(* Logix 5000 project; controller R400_500_XLS vendor 1 type 14 code 216 rev 31.11; software revision 31.01; part 13 of 32 *)
(* tags used below, declared in another part *)
   Alarm : SINT;   // Wait 3 seconds
   AlarmMuted : BOOL;
   Chem_Pump : UDT_CHEM_PUMP[4];   // Chemical Pump flow rate
   ChPumpRunningTime : REAL;
   Inj_Cond : SINT;   // Conductivity injection based steps
   Inj_Time : SINT;   // Time based chemical injection steps
   M : DINT[5];   // Memory Bits
   NeutralizantPump : SINT;
   NeutralizationInjTime : DINT;
   NeutralizationRecircTime : DINT;
   OneShot : DINT[1];
   Run : DINT;
   Service : DINT[2];   // Unused Service Mode Memory Bit
   Supervisor : DINT;
   Tmr : TIMER[107];
   VolumeInjected_ML : REAL;
   VolumeNeutralizer : REAL;
   washerMode : SINT;   // Washer Mode Flag 0 -> Ready; 1 -> Supervisor; 2 -> Service; 3 -> Run.
   WshExcBuffer : UDT_WASH;
   Current_Screen : DINT;
   Doors_Check : DINT;
   NumInput : UDT_NUMERIC_INPUT[65];   // Numeric input
   NumInputReal : UDT_NUMERIC_INPUT_REAL[17];
   Q_Chm_1 : BOOL;   // Chemical pump #1
   Q_Chm_2 : BOOL;   // Chemical pump #2
   Q_Chm_3 : BOOL;   // Chemical pump #3
   Q_Chm_4 : BOOL;   // Chemical pump #4
   Screen_Ctrl : DINT;   // PLC Screen Request
   SelChemNeutralizer : UDT_SELECTOR[5];
   SelChemNeutralizerESign : UDT_SELECTOR[5];
   Selector : UDT_SELECTOR[25];   // Piloted list selector
   Tpb : DINT[11];
   udtAudibleAlarmMode : UDT_SELECTOR;
   Unit : Hrdwre;   // Unit Configuration
(* MainProgram, continued *)

ROUTINE SPV_18_AUDIBLE_ALARM_OP_MODE   (* ladder *)
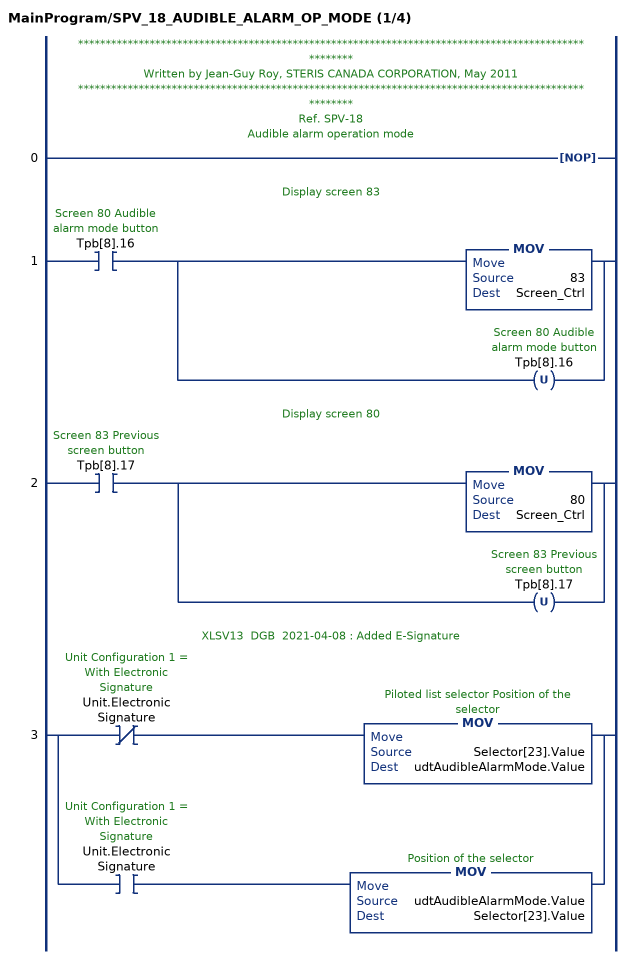
   // ****************************************************************************************************
   // Written by Jean-Guy Roy, STERIS CANADA CORPORATION, May 2011
   // ****************************************************************************************************
   // Ref. SPV-18
   // Audible alarm operation mode
   0: NOP();
   // Display screen 83
   1: XIC(Tpb[8].16)[MOV(83,Screen_Ctrl) ,OTU(Tpb[8].16) ];
   // Display screen 80
   2: XIC(Tpb[8].17)[MOV(80,Screen_Ctrl) ,OTU(Tpb[8].17) ];
   // XLSV13  DGB  2021-04-08 : Added E-Signature
   3: [XIO(Unit.ElectronicSignature) MOV(Selector[23].Value,udtAudibleAlarmMode.Value) ,XIC(Unit.ElectronicSignature) MOV(udtAudibleAlarmMode.Value,Selector[23].Value) ];
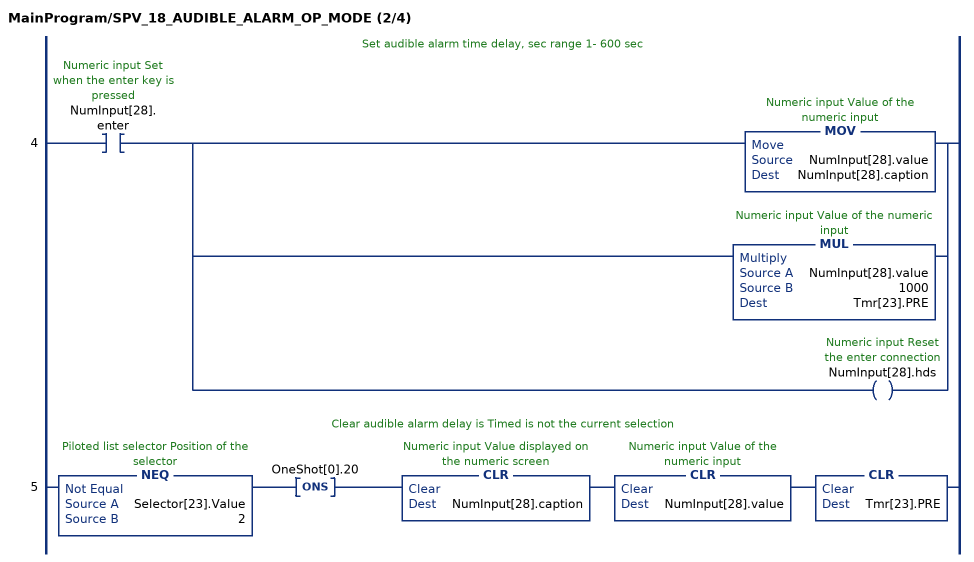
   // Set audible alarm time delay, sec range 1- 600 sec
   4: XIC(NumInput[28].enter)[MOV(NumInput[28].value,NumInput[28].caption) ,MUL(NumInput[28].value,1000,Tmr[23].PRE) ,OTE(NumInput[28].hds) ];
   // Clear audible alarm delay is Timed is not the current selection
   5: NEQ(Selector[23].Value,2)ONS(OneShot[0].20)CLR(NumInput[28].caption)CLR(NumInput[28].value)CLR(Tmr[23].PRE);
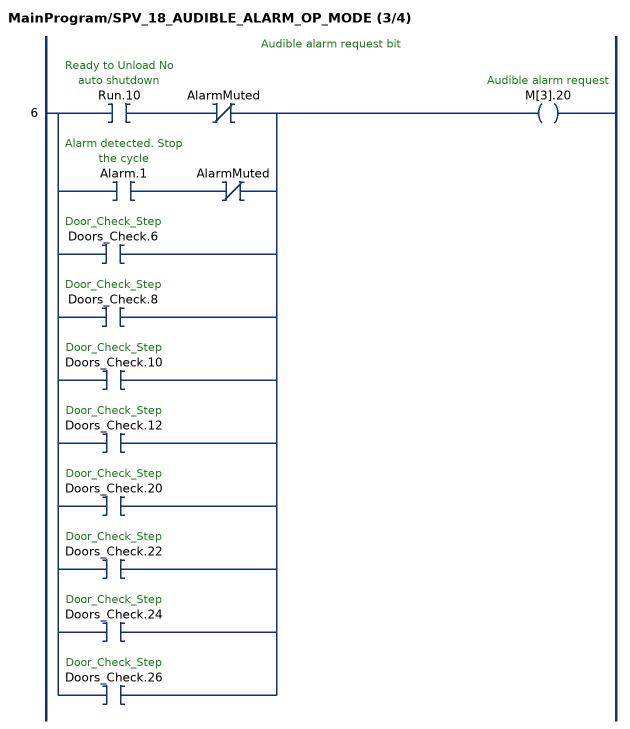
   // Audible alarm request bit
   6: [XIC(Run.10) XIO(AlarmMuted) ,XIC(Alarm.1) XIO(AlarmMuted) ,XIC(Doors_Check.6) ,XIC(Doors_Check.8) ,XIC(Doors_Check.10) ,XIC(Doors_Check.12) ,XIC(Doors_Check.20) ,XIC(Doors_Check.22) ,XIC(Doors_Check.24) ,XIC(Doors_Check.26) ]OTE(M[3].20);
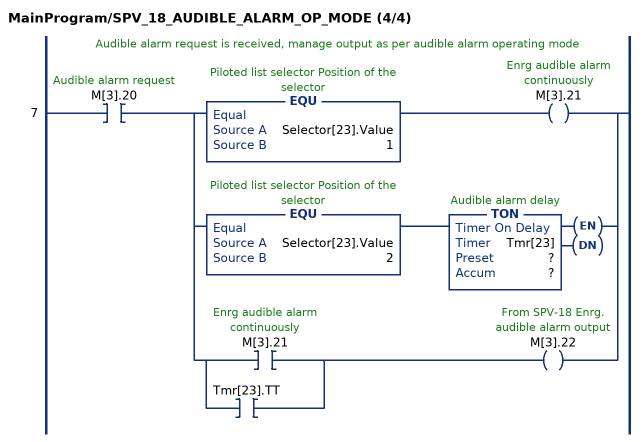
   // Audible alarm request is received, manage output as per audible alarm operating mode
   7: XIC(M[3].20)[EQU(Selector[23].Value,1) OTE(M[3].21) ,EQU(Selector[23].Value,2) TON(Tmr[23],?,?) ,[XIC(M[3].21) ,XIC(Tmr[23].TT) ] OTE(M[3].22) ];
END_ROUTINE

ROUTINE SPV_1_SUPERVISOR_ACCESS   (* ladder *)
// Screen Control routine
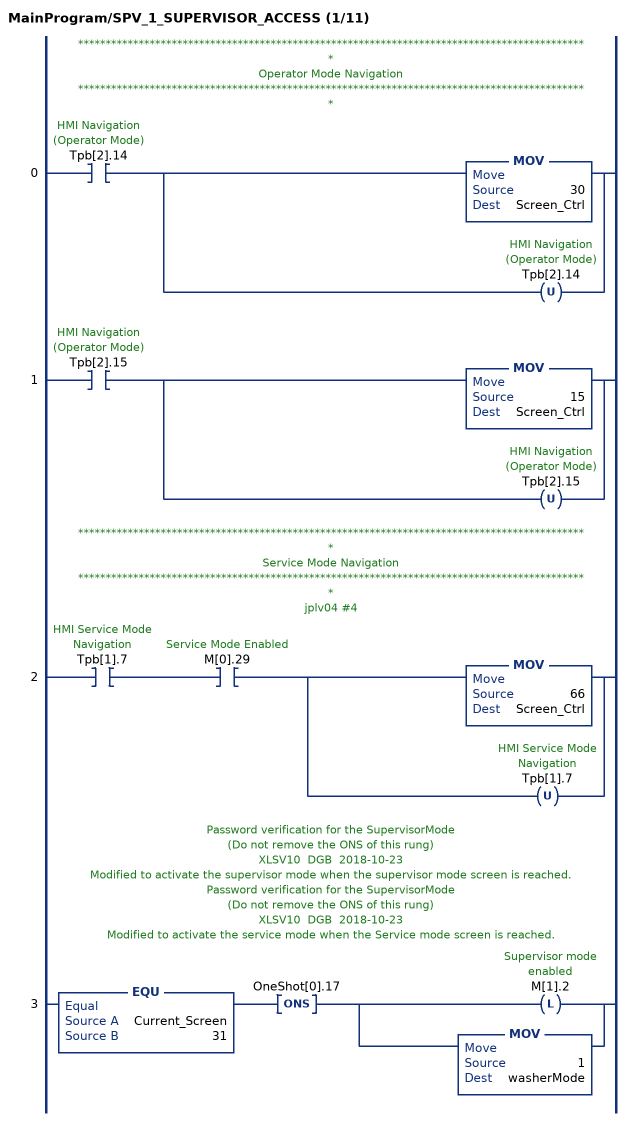
   // *********************************************************************************************
   // Operator Mode Navigation
   // *********************************************************************************************
   0: XIC(Tpb[2].14)[MOV(30,Screen_Ctrl) ,OTU(Tpb[2].14) ];
   1: XIC(Tpb[2].15)[MOV(15,Screen_Ctrl) ,OTU(Tpb[2].15) ];
   // *********************************************************************************************
   // Service Mode Navigation
   // *********************************************************************************************
   // jplv04 #4
   2: XIC(Tpb[1].7)XIC(M[0].29)[MOV(66,Screen_Ctrl) ,OTU(Tpb[1].7) ];
   // Password verification for the SupervisorMode
   // (Do not remove the ONS of this rung)
   // XLSV10  DGB  2018-10-23
   // Modified to activate the supervisor mode when the supervisor mode screen is reached.
   // Password verification for the SupervisorMode
   // (Do not remove the ONS of this rung)
   // XLSV10  DGB  2018-10-23
   // Modified to activate the service mode when the Service mode screen is reached.
   3: EQU(Current_Screen,31)ONS(OneShot[0].17)[OTL(M[1].2) ,MOV(1,washerMode) ];
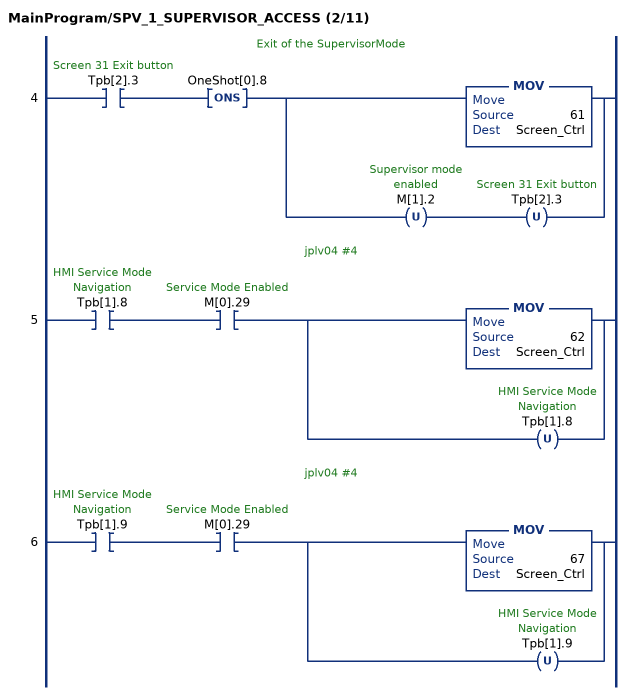
   // Exit of the SupervisorMode
   4: XIC(Tpb[2].3)ONS(OneShot[0].8)[MOV(61,Screen_Ctrl) ,OTU(M[1].2) OTU(Tpb[2].3) ];
   // jplv04 #4
   5: XIC(Tpb[1].8)XIC(M[0].29)[MOV(62,Screen_Ctrl) ,OTU(Tpb[1].8) ];
   // jplv04 #4
   6: XIC(Tpb[1].9)XIC(M[0].29)[MOV(67,Screen_Ctrl) ,OTU(Tpb[1].9) ];
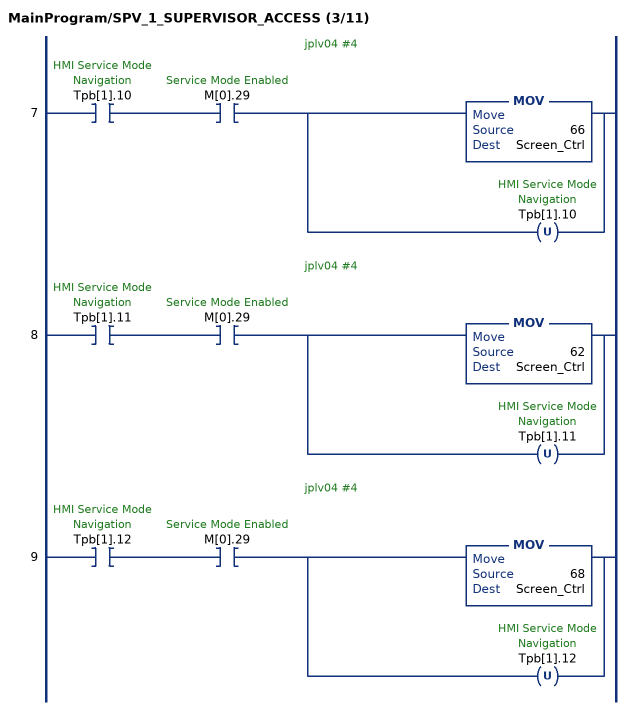
   // jplv04 #4
   7: XIC(Tpb[1].10)XIC(M[0].29)[MOV(66,Screen_Ctrl) ,OTU(Tpb[1].10) ];
   // jplv04 #4
   8: XIC(Tpb[1].11)XIC(M[0].29)[MOV(62,Screen_Ctrl) ,OTU(Tpb[1].11) ];
   // jplv04 #4
   9: XIC(Tpb[1].12)XIC(M[0].29)[MOV(68,Screen_Ctrl) ,OTU(Tpb[1].12) ];
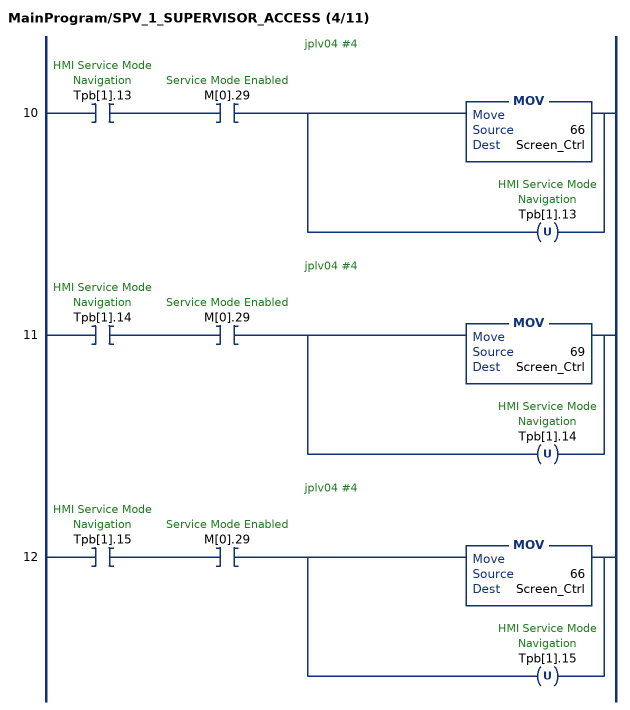
   // jplv04 #4
   10: XIC(Tpb[1].13)XIC(M[0].29)[MOV(66,Screen_Ctrl) ,OTU(Tpb[1].13) ];
   // jplv04 #4
   11: XIC(Tpb[1].14)XIC(M[0].29)[MOV(69,Screen_Ctrl) ,OTU(Tpb[1].14) ];
   // jplv04 #4
   12: XIC(Tpb[1].15)XIC(M[0].29)[MOV(66,Screen_Ctrl) ,OTU(Tpb[1].15) ];
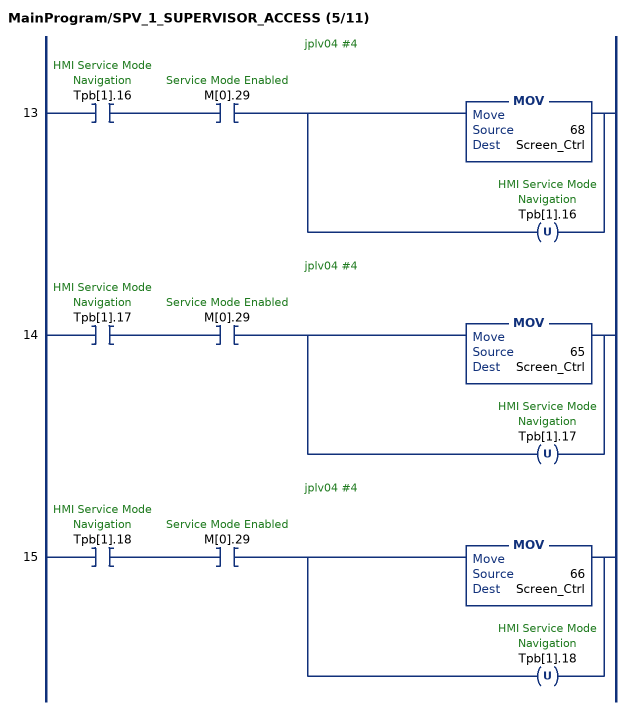
   // jplv04 #4
   13: XIC(Tpb[1].16)XIC(M[0].29)[MOV(68,Screen_Ctrl) ,OTU(Tpb[1].16) ];
   // jplv04 #4
   14: XIC(Tpb[1].17)XIC(M[0].29)[MOV(65,Screen_Ctrl) ,OTU(Tpb[1].17) ];
   // jplv04 #4
   15: XIC(Tpb[1].18)XIC(M[0].29)[MOV(66,Screen_Ctrl) ,OTU(Tpb[1].18) ];
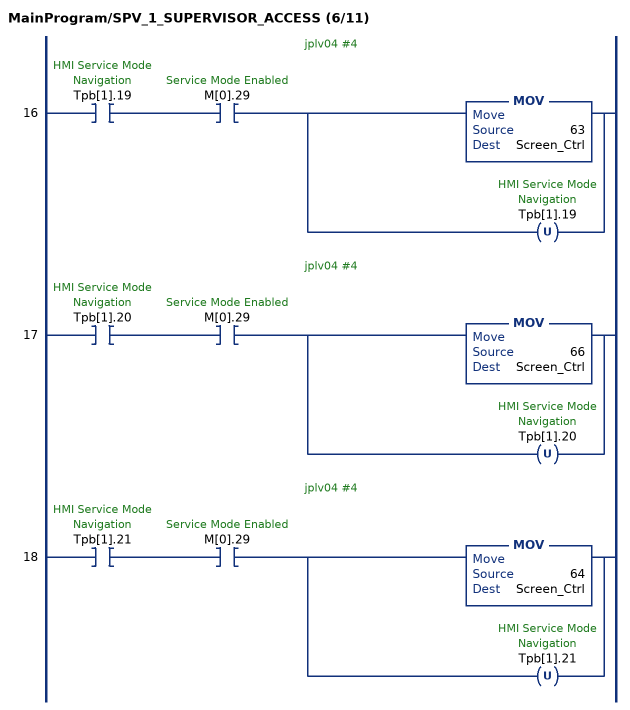
   // jplv04 #4
   16: XIC(Tpb[1].19)XIC(M[0].29)[MOV(63,Screen_Ctrl) ,OTU(Tpb[1].19) ];
   // jplv04 #4
   17: XIC(Tpb[1].20)XIC(M[0].29)[MOV(66,Screen_Ctrl) ,OTU(Tpb[1].20) ];
   // jplv04 #4
   18: XIC(Tpb[1].21)XIC(M[0].29)[MOV(64,Screen_Ctrl) ,OTU(Tpb[1].21) ];
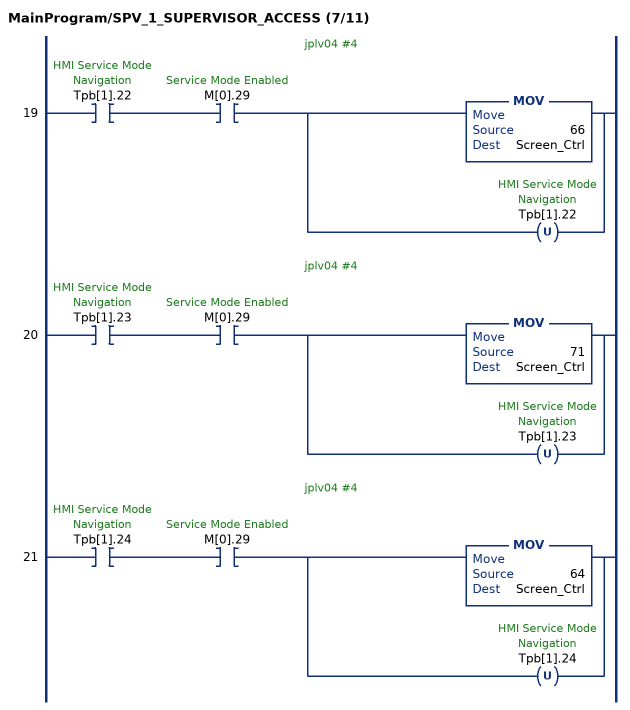
   // jplv04 #4
   19: XIC(Tpb[1].22)XIC(M[0].29)[MOV(66,Screen_Ctrl) ,OTU(Tpb[1].22) ];
   // jplv04 #4
   20: XIC(Tpb[1].23)XIC(M[0].29)[MOV(71,Screen_Ctrl) ,OTU(Tpb[1].23) ];
   // jplv04 #4
   21: XIC(Tpb[1].24)XIC(M[0].29)[MOV(64,Screen_Ctrl) ,OTU(Tpb[1].24) ];
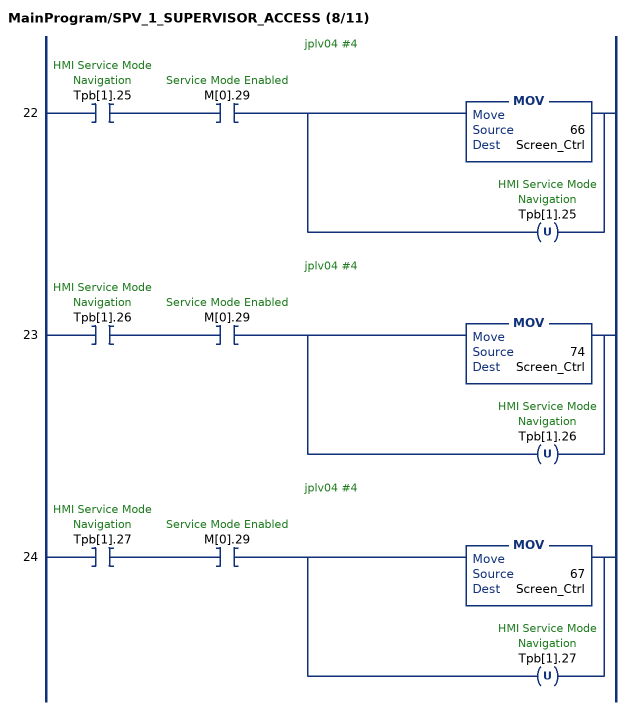
   // jplv04 #4
   22: XIC(Tpb[1].25)XIC(M[0].29)[MOV(66,Screen_Ctrl) ,OTU(Tpb[1].25) ];
   // jplv04 #4
   23: XIC(Tpb[1].26)XIC(M[0].29)[MOV(74,Screen_Ctrl) ,OTU(Tpb[1].26) ];
   // jplv04 #4
   24: XIC(Tpb[1].27)XIC(M[0].29)[MOV(67,Screen_Ctrl) ,OTU(Tpb[1].27) ];
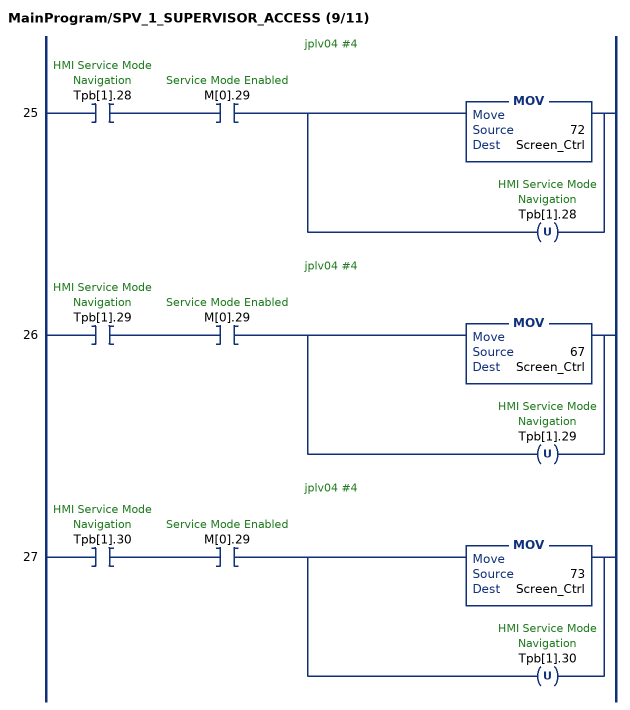
   // jplv04 #4
   25: XIC(Tpb[1].28)XIC(M[0].29)[MOV(72,Screen_Ctrl) ,OTU(Tpb[1].28) ];
   // jplv04 #4
   26: XIC(Tpb[1].29)XIC(M[0].29)[MOV(67,Screen_Ctrl) ,OTU(Tpb[1].29) ];
   // jplv04 #4
   27: XIC(Tpb[1].30)XIC(M[0].29)[MOV(73,Screen_Ctrl) ,OTU(Tpb[1].30) ];
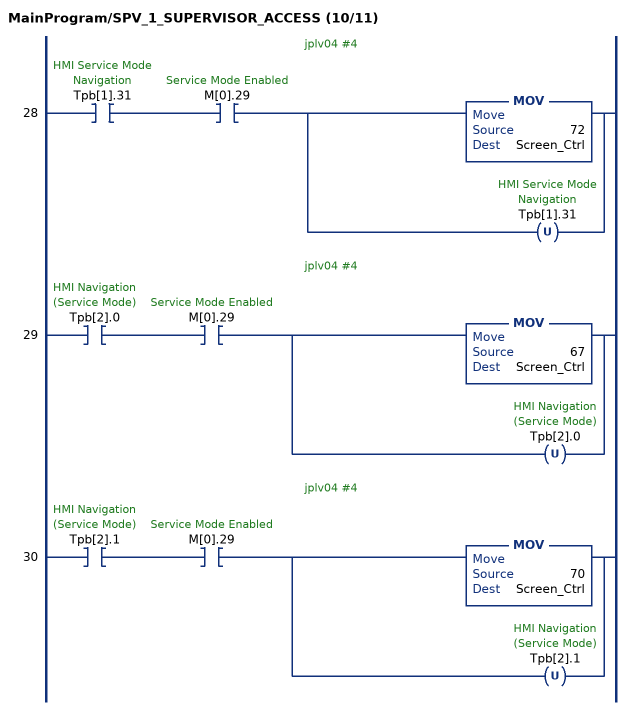
   // jplv04 #4
   28: XIC(Tpb[1].31)XIC(M[0].29)[MOV(72,Screen_Ctrl) ,OTU(Tpb[1].31) ];
   // jplv04 #4
   29: XIC(Tpb[2].0)XIC(M[0].29)[MOV(67,Screen_Ctrl) ,OTU(Tpb[2].0) ];
   // jplv04 #4
   30: XIC(Tpb[2].1)XIC(M[0].29)[MOV(70,Screen_Ctrl) ,OTU(Tpb[2].1) ];
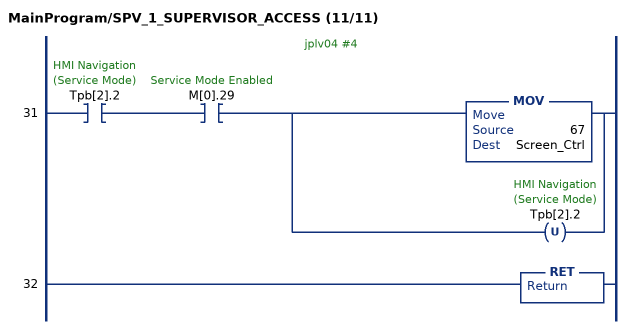
   // jplv04 #4
   31: XIC(Tpb[2].2)XIC(M[0].29)[MOV(67,Screen_Ctrl) ,OTU(Tpb[2].2) ];
   32: RET();
END_ROUTINE

ROUTINE SPV_21_UNITS   (* ladder *)
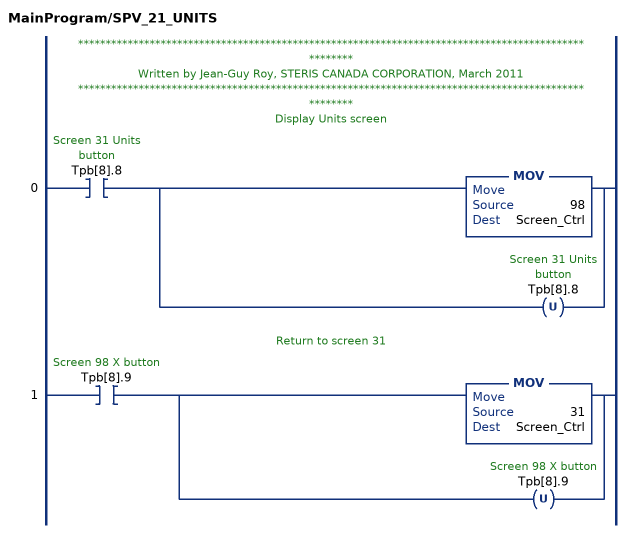
   // ****************************************************************************************************
   // Written by Jean-Guy Roy, STERIS CANADA CORPORATION, March 2011
   // ****************************************************************************************************
   // Display Units screen
   0: XIC(Tpb[8].8)[MOV(98,Screen_Ctrl) ,OTU(Tpb[8].8) ];
   // Return to screen 31
   1: XIC(Tpb[8].9)[MOV(31,Screen_Ctrl) ,OTU(Tpb[8].9) ];
END_ROUTINE

ROUTINE SPV_22_WSH_35_NEUTRALIZATION   (* ladder *)
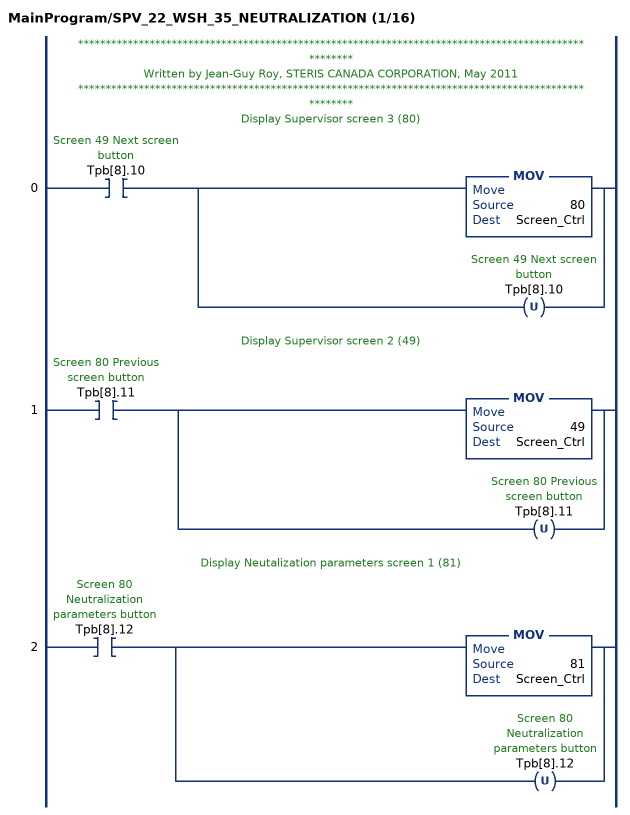
   // ****************************************************************************************************
   // Written by Jean-Guy Roy, STERIS CANADA CORPORATION, May 2011
   // ****************************************************************************************************
   // Display Supervisor screen 3 (80)
   0: XIC(Tpb[8].10)[MOV(80,Screen_Ctrl) ,OTU(Tpb[8].10) ];
   // Display Supervisor screen 2 (49)
   1: XIC(Tpb[8].11)[MOV(49,Screen_Ctrl) ,OTU(Tpb[8].11) ];
   // Display Neutalization parameters screen 1 (81)
   2: XIC(Tpb[8].12)[MOV(81,Screen_Ctrl) ,OTU(Tpb[8].12) ];
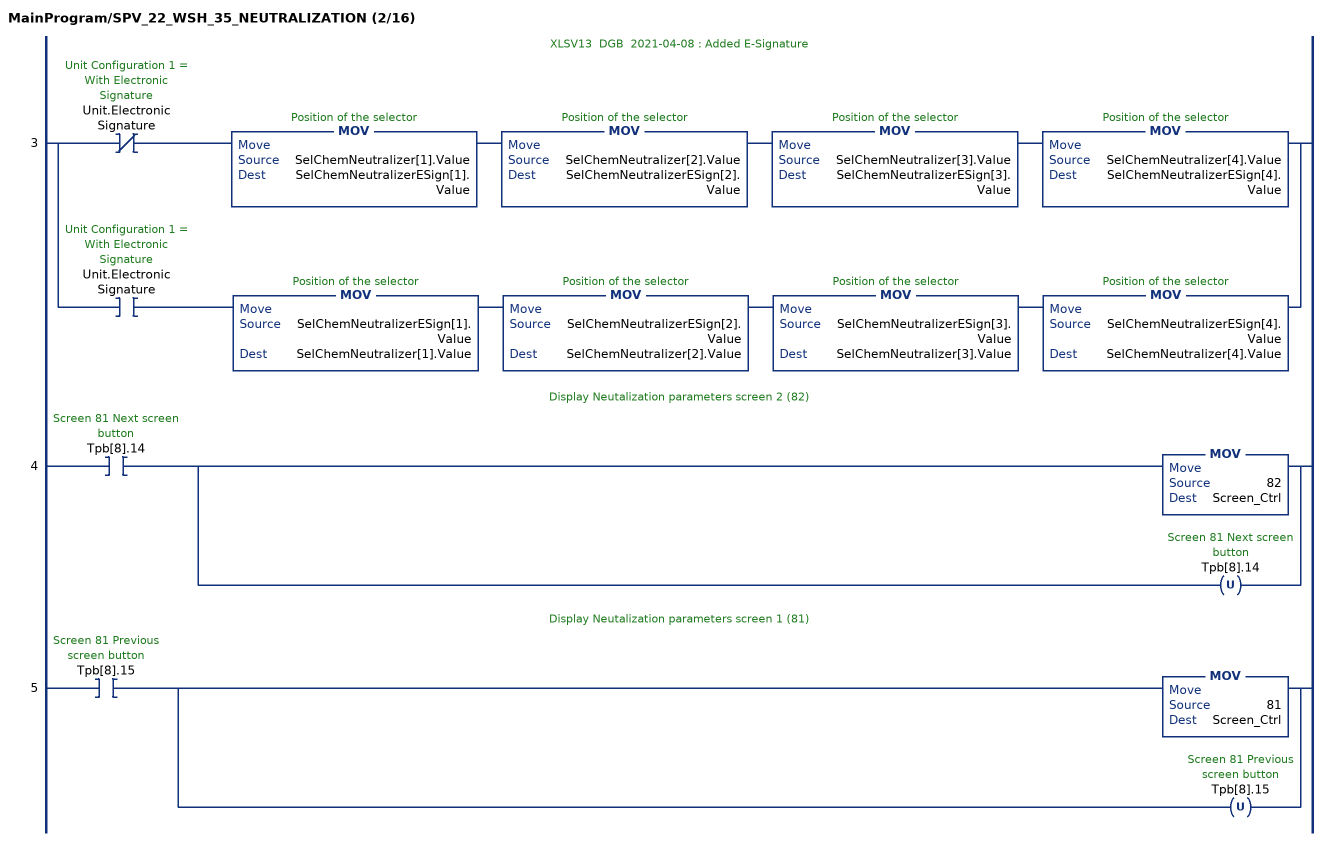
   // XLSV13  DGB  2021-04-08 : Added E-Signature
   3: [XIO(Unit.ElectronicSignature) MOV(SelChemNeutralizer[1].Value,SelChemNeutralizerESign[1].Value) MOV(SelChemNeutralizer[2].Value,SelChemNeutralizerESign[2].Value) MOV(SelChemNeutralizer[3].Value,SelChemNeutralizerESign[3].Value) MOV(SelChemNeutralizer[4].Value,SelChemNeutralizerESign[4].Value) ,XIC(Unit.ElectronicSignature) MOV(SelChemNeutralizerESign[1].Value,SelChemNeutralizer[1].Value) MOV(SelChemNeutralizerESign[2].Value,SelChemNeutralizer[2].Value) MOV(SelChemNeutralizerESign[3].Value,SelChemNeutralizer[3].Value) MOV(SelChemNeutralizerESign[4].Value,SelChemNeutralizer[4].Value) ];
   // Display Neutalization parameters screen 2 (82)
   4: XIC(Tpb[8].14)[MOV(82,Screen_Ctrl) ,OTU(Tpb[8].14) ];
   // Display Neutalization parameters screen 1 (81)
   5: XIC(Tpb[8].15)[MOV(81,Screen_Ctrl) ,OTU(Tpb[8].15) ];
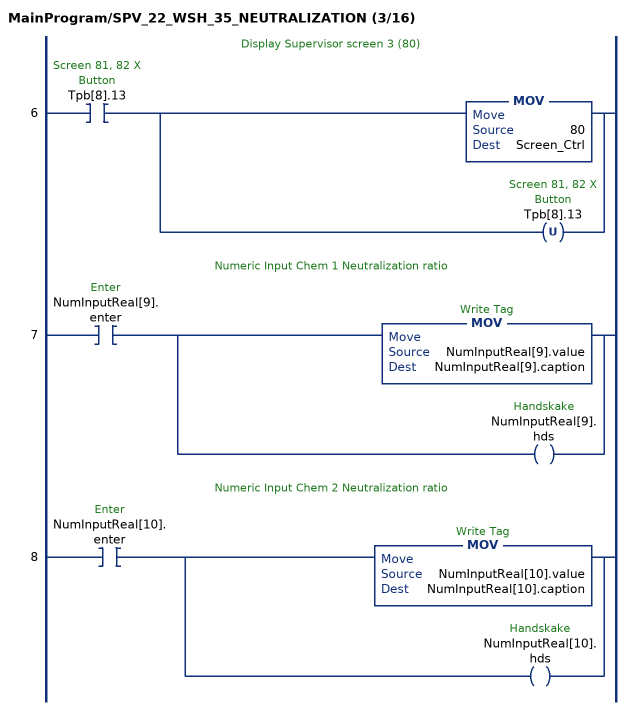
   // Display Supervisor screen 3 (80)
   6: XIC(Tpb[8].13)[MOV(80,Screen_Ctrl) ,OTU(Tpb[8].13) ];
   // Numeric Input Chem 1 Neutralization ratio
   7: XIC(NumInputReal[9].enter)[MOV(NumInputReal[9].value,NumInputReal[9].caption) ,OTE(NumInputReal[9].hds) ];
   // Numeric Input Chem 2 Neutralization ratio
   8: XIC(NumInputReal[10].enter)[MOV(NumInputReal[10].value,NumInputReal[10].caption) ,OTE(NumInputReal[10].hds) ];
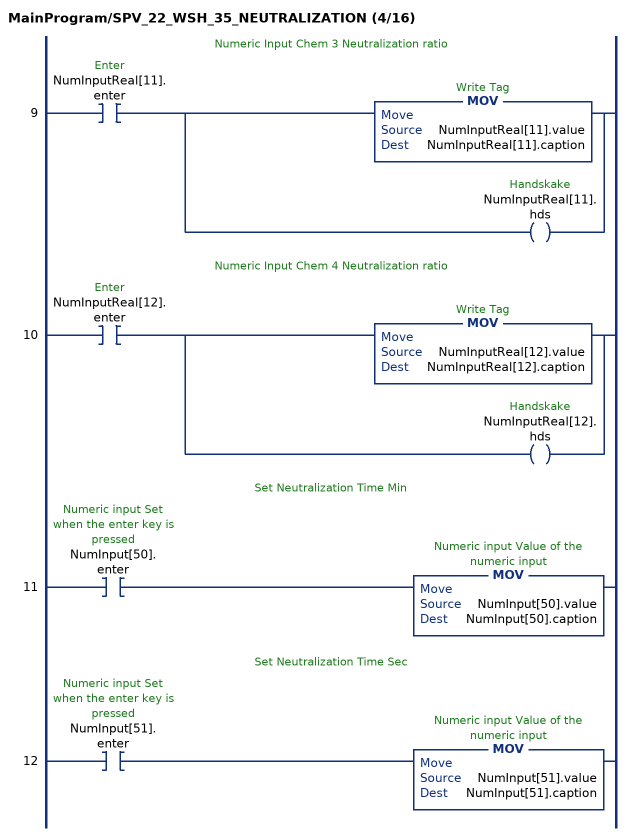
   // Numeric Input Chem 3 Neutralization ratio
   9: XIC(NumInputReal[11].enter)[MOV(NumInputReal[11].value,NumInputReal[11].caption) ,OTE(NumInputReal[11].hds) ];
   // Numeric Input Chem 4 Neutralization ratio
   10: XIC(NumInputReal[12].enter)[MOV(NumInputReal[12].value,NumInputReal[12].caption) ,OTE(NumInputReal[12].hds) ];
   // Set Neutralization Time Min
   11: XIC(NumInput[50].enter)MOV(NumInput[50].value,NumInput[50].caption);
   // Set Neutralization Time Sec
   12: XIC(NumInput[51].enter)MOV(NumInput[51].value,NumInput[51].caption);
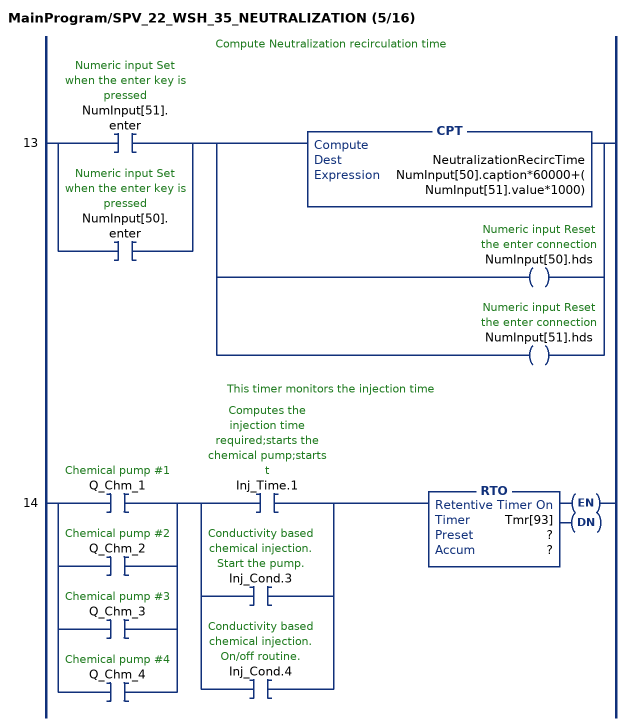
   // Compute Neutralization recirculation time
   13: [XIC(NumInput[51].enter) ,XIC(NumInput[50].enter) ][CPT(NeutralizationRecircTime,NumInput[50].caption*60000+(NumInput[51].value*1000)) ,OTE(NumInput[50].hds) ,OTE(NumInput[51].hds) ];
   // This timer monitors the injection time
   14: [XIC(Q_Chm_1) ,XIC(Q_Chm_2) ,XIC(Q_Chm_3) ,XIC(Q_Chm_4) ][XIC(Inj_Time.1) ,XIC(Inj_Cond.3) ,XIC(Inj_Cond.4) ]RTO(Tmr[93],?,?);
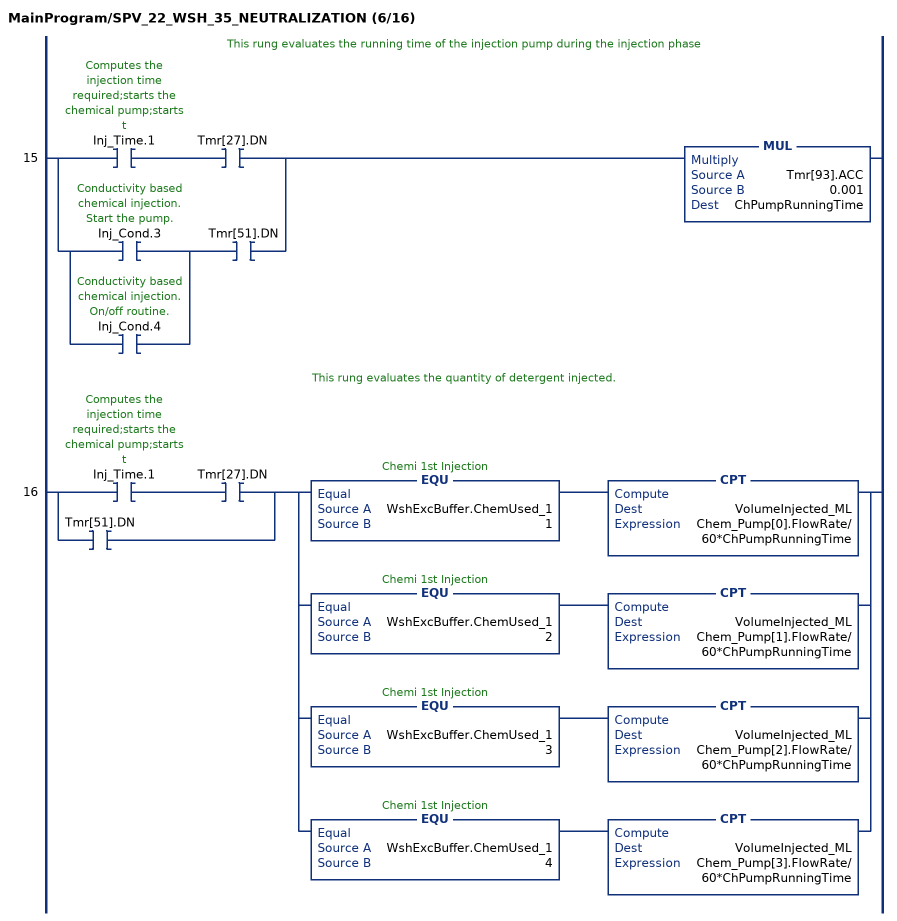
   // This rung evaluates the running time of the injection pump during the injection phase
   15: [XIC(Inj_Time.1) XIC(Tmr[27].DN) ,[XIC(Inj_Cond.3) ,XIC(Inj_Cond.4) ] XIC(Tmr[51].DN) ]MUL(Tmr[93].ACC,0.001,ChPumpRunningTime);
   // This rung evaluates the quantity of detergent injected.
   16: [XIC(Inj_Time.1) XIC(Tmr[27].DN) ,XIC(Tmr[51].DN) ][EQU(WshExcBuffer.ChemUsed_1,1) CPT(VolumeInjected_ML,Chem_Pump[0].FlowRate/60*ChPumpRunningTime) ,EQU(WshExcBuffer.ChemUsed_1,2) CPT(VolumeInjected_ML,Chem_Pump[1].FlowRate/60*ChPumpRunningTime) ,EQU(WshExcBuffer.ChemUsed_1,3) CPT(VolumeInjected_ML,Chem_Pump[2].FlowRate/60*ChPumpRunningTime) ,EQU(WshExcBuffer.ChemUsed_1,4) CPT(VolumeInjected_ML,Chem_Pump[3].FlowRate/60*ChPumpRunningTime) ];
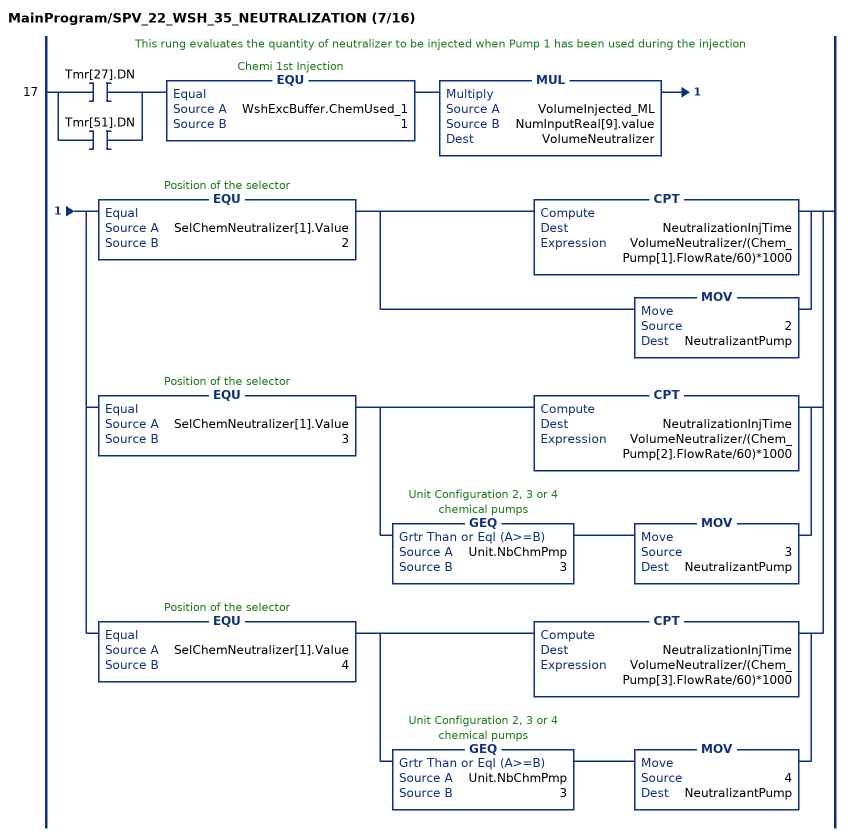
   // This rung evaluates the quantity of neutralizer to be injected when Pump 1 has been used during the injection
   17: [XIC(Tmr[27].DN) ,XIC(Tmr[51].DN) ]EQU(WshExcBuffer.ChemUsed_1,1)MUL(VolumeInjected_ML,NumInputReal[9].value,VolumeNeutralizer)[EQU(SelChemNeutralizer[1].Value,2) [CPT(NeutralizationInjTime,VolumeNeutralizer/(Chem_Pump[1].FlowRate/60)*1000) ,MOV(2,NeutralizantPump) ] ,EQU(SelChemNeutralizer[1].Value,3) [CPT(NeutralizationInjTime,VolumeNeutralizer/(Chem_Pump[2].FlowRate/60)*1000) ,GEQ(Unit.NbChmPmp,3) MOV(3,NeutralizantPump) ] ,EQU(SelChemNeutralizer[1].Value,4) [CPT(NeutralizationInjTime,VolumeNeutralizer/(Chem_Pump[3].FlowRate/60)*1000) ,GEQ(Unit.NbChmPmp,3) MOV(4,NeutralizantPump) ] ];
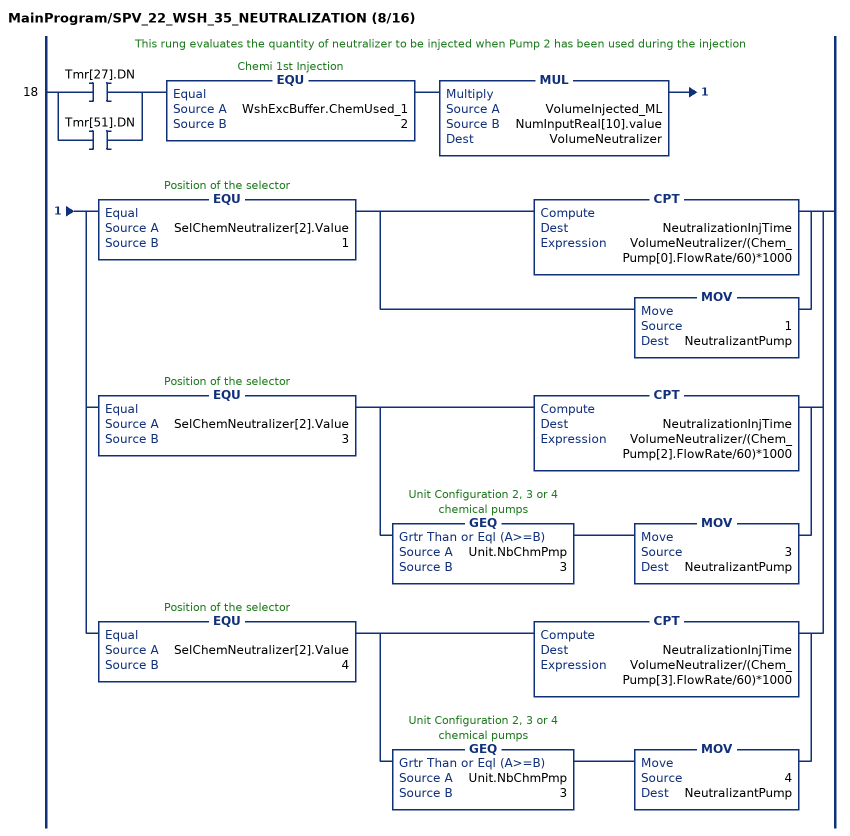
   // This rung evaluates the quantity of neutralizer to be injected when Pump 2 has been used during the injection
   18: [XIC(Tmr[27].DN) ,XIC(Tmr[51].DN) ]EQU(WshExcBuffer.ChemUsed_1,2)MUL(VolumeInjected_ML,NumInputReal[10].value,VolumeNeutralizer)[EQU(SelChemNeutralizer[2].Value,1) [CPT(NeutralizationInjTime,VolumeNeutralizer/(Chem_Pump[0].FlowRate/60)*1000) ,MOV(1,NeutralizantPump) ] ,EQU(SelChemNeutralizer[2].Value,3) [CPT(NeutralizationInjTime,VolumeNeutralizer/(Chem_Pump[2].FlowRate/60)*1000) ,GEQ(Unit.NbChmPmp,3) MOV(3,NeutralizantPump) ] ,EQU(SelChemNeutralizer[2].Value,4) [CPT(NeutralizationInjTime,VolumeNeutralizer/(Chem_Pump[3].FlowRate/60)*1000) ,GEQ(Unit.NbChmPmp,3) MOV(4,NeutralizantPump) ] ];
